(* Schneider Machine Expert - Basic project modbus_full_pin_write, file version 3.0.0.0 *)
(* ProjectInformations: Name=New project *)

HARDWARE
  Cpu 0: TM200CE40T
  EthernetConfiguration: NetworkName=M200, IpAllocationMode=FixedAddress, IpAddress=0.0.0.0, SubnetMask=0.0.0.0
  SerialLineConfiguration: Baud=Baud19200, Parity=ParityEven, DataBits=DataBits8, StopBits=StopBits1, PhysicalMedium=PhysicalMediumRs485, TransmissionMode=TransmissionModeModbusRtu, SlaveId=1, Addressing=MasterAddressing
  MastTask: UsePeriodScanMode=false, PeriodScan=100
  FastTask: Period=255
  CpuBehavior: StartingMode=StartAsPreviousState, AutoSaveRamOnEeprom=true, WatchdogPeriod=250

SYMBOLS  (address, symbol, comment, settings)
  %WRITE_VAR0   [Link(Value(FBComLinkParameterEnums=SerialLine1)), RemoteDeviceId(Value(int=1)), Timeout(Value(int=100)), ObjType(Value(FBComObjTypeParameterEnums=Q)), FirstObj(Value(int=73)), Quantity(Value(int=17)), IndexData(Value(int=240))]

POU Generated C++ - EXPERIMENTAL
  (* SectionNumber=0 *)

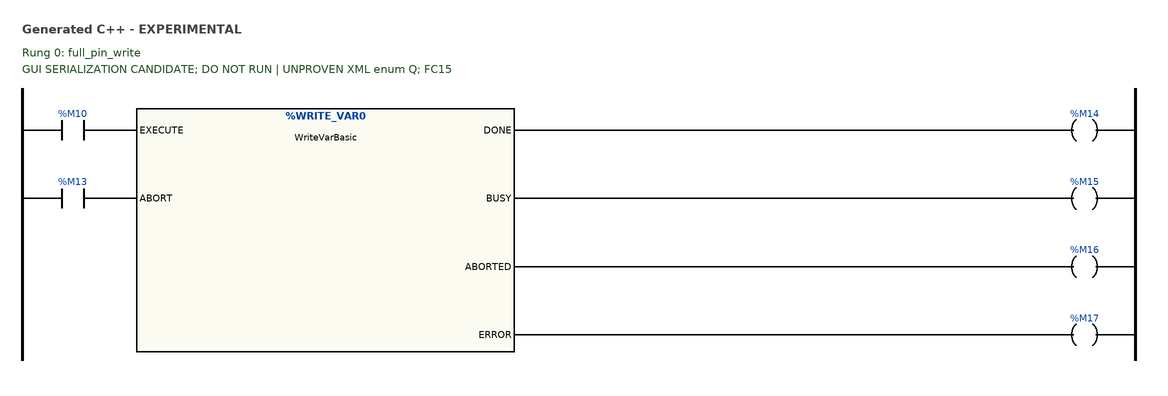

// Rung 0: full_pin_write
// GUI SERIALIZATION CANDIDATE; DO NOT RUN | UNPROVEN XML enum Q; FC15
  BLK %WRITE_VAR0
  LD %M10
  EXECUTE
  LD %M13
  ABORT
  OUT_BLK
  LD DONE
  ST %M14
  LD BUSY
  ST %M15
  LD ABORTED
  ST %M16
  LD ERROR
  ST %M17
  END_BLK
  // as ST:
  //   %WRITE_VAR0(EXECUTE := %M10, ABORT := %M13);
  //   %M14 := %WRITE_VAR0.DONE;
  //   %M15 := %WRITE_VAR0.BUSY;
  //   %M16 := %WRITE_VAR0.ABORTED;
  //   %M17 := %WRITE_VAR0.ERROR;
